{attribute 'pack_mode' := '1'} 
// ------------------------------------------------------------------------- 
//  SRCI Robot Library                                                
// ------------------------------------------------------------------------- 
//                                                                           
//  Object:      TelegramPlcToRobCyclicData                                       
//  Author:      Thorsten Brach                                                
//  Date:        2024-11-30
//
//  Description:                                              
//   
//                                                                           
//  Copyright: 
//    (C) 2024 Thorsten Brach. All rights reserved                                                                                                                                            
//             Licensed under the MIT License.
//                                                                           
//  Disclaimer:                                                                           
//    This project is provided without any guarantee and can be used for   
//    private and commercial purposes. Any use is at the user’s 
//    own risk and responsibility.
//
// -------------------------------------------------------------------------
TYPE TelegramPlcToRobCyclicData :
STRUCT
  /// Current Tool
  ToolNo  : BYTE;
  /// Current Frame
  FrameNo : BYTE;      
END_STRUCT
END_TYPE

{attribute 'pack_mode' := '1'} 
// ------------------------------------------------------------------------- 
//  SRCI Robot Library                                                
// ------------------------------------------------------------------------- 
//                                                                           
//  Object:      TelegramPlcToRobCyclicOptionalCartesianPos                                       
//  Author:      Thorsten Brach                                                
//  Date:        2024-06-01
//
//  Description:                                              
//   
//                                                                           
//  Copyright: 
//    (C) 2024 Thorsten Brach. All rights reserved                                                                                                                                            
//             Licensed under the MIT License.
//                                                                           
//  Disclaimer:                                                                           
//    This project is provided without any guarantee and can be used for   
//    private and commercial purposes. Any use is at the user’s 
//    own risk and responsibility.
//
// -------------------------------------------------------------------------
TYPE TelegramPlcToRobCyclicOptionalCartesianPosition :
STRUCT
  /// TCP Position on the X-Axis
  X           : REAL;
  /// TCP Position on the Y-Axis
  Y           : REAL;
  /// TCP Position on the Z-Axis
  Z           : REAL;
  /// Rotation around the X-Axis (RX)
  Rx          : REAL;
  /// Rotation around the Y-Axis (RY)
  Ry          : REAL;
  /// Rotation around the Z-Axis (RZ)
  Rz          : REAL;
  /// Configuration
  Config      : WORD;
  /// Turns of J1 and J2
  Turns_J2_J1 : BYTE;
  /// Turns of J3 and J4
  Turns_J4_J3 : BYTE;
  /// Turns of J6 and J5
  Turns_J6_J5 : BYTE;
  /// Turns of E1
  Turns_E1    : BYTE;
  /// Position of first external axis
  E1          : REAL;
END_STRUCT
END_TYPE

{attribute 'pack_mode' := '1'} 
// ------------------------------------------------------------------------- 
//  SRCI Robot Library                                                
// ------------------------------------------------------------------------- 
//                                                                           
//  Object:      TelegramPlcToRobCyclicOptionalCartesianPositionExt                                       
//  Author:      Thorsten Brach                                                
//  Date:        2024-06-01
//
//  Description:                                              
//   
//                                                                           
//  Copyright: 
//    (C) 2024 Thorsten Brach. All rights reserved                                                                                                                                            
//             Licensed under the MIT License.
//                                                                           
//  Disclaimer:                                                                           
//    This project is provided without any guarantee and can be used for   
//    private and commercial purposes. Any use is at the user’s 
//    own risk and responsibility.
//
// -------------------------------------------------------------------------
TYPE TelegramPlcToRobCyclicOptionalCartesianPositionExt :
STRUCT
  /// Position of second external axis
  E2 : REAL;
  /// Position of third external axis
  E3 : REAL;
  /// Position of fourth external axis
  E4 : REAL;
  /// Position of fifth external axis
  E5 : REAL;
  /// Position of sixth external axis
  E6 : REAL;    
END_STRUCT
END_TYPE

{attribute 'pack_mode' := '1'} 
// ------------------------------------------------------------------------- 
//  SRCI Robot Library                                                
// ------------------------------------------------------------------------- 
//                                                                           
//  Object:      TelegramPlcToRobCyclicOptionalCurrent                                       
//  Author:      Thorsten Brach                                                
//  Date:        2024-06-01
//
//  Description:                                              
//   
//                                                                           
//  Copyright: 
//    (C) 2024 Thorsten Brach. All rights reserved                                                                                                                                            
//             Licensed under the MIT License.
//                                                                           
//  Disclaimer:                                                                           
//    This project is provided without any guarantee and can be used for   
//    private and commercial purposes. Any use is at the user’s 
//    own risk and responsibility.
//
// -------------------------------------------------------------------------
TYPE TelegramPlcToRobCyclicOptionalCurrent :
STRUCT
  /// Current of first joint of the robot
  J1 : REAL;
  /// Current of second joint of the robot
  J2 : REAL;
  /// Current of third joint of the robot
  J3 : REAL;
  /// Current of fourth joint of the robot
  J4 : REAL;
  /// Current of fifth joint of the robot
  J5 : REAL;
  /// Current of sixth joint of the robot
  J6 : REAL;  
END_STRUCT
END_TYPE

{attribute 'pack_mode' := '1'} 
// ------------------------------------------------------------------------- 
//  SRCI Robot Library                                                
// ------------------------------------------------------------------------- 
//                                                                           
//  Object:      TelegramPlcToRobCyclicOptionalCurrentExt                                       
//  Author:      Thorsten Brach                                                
//  Date:        2024-06-01
//
//  Description:                                              
//   
//                                                                           
//  Copyright: 
//    (C) 2024 Thorsten Brach. All rights reserved                                                                                                                                            
//             Licensed under the MIT License.
//                                                                           
//  Disclaimer:                                                                           
//    This project is provided without any guarantee and can be used for   
//    private and commercial purposes. Any use is at the user’s 
//    own risk and responsibility.
//
// -------------------------------------------------------------------------
TYPE TelegramPlcToRobCyclicOptionalCurrentExt :
STRUCT
  /// Current of first external joint of the robot
  E1 : REAL;
  /// Current of second external axis
  E2: REAL;
  /// Current of third external axis
  E3: REAL;
  /// Current of fourth external axis
  E4: REAL;
  /// Current of fifth external axis
  E5: REAL;
  /// Current of sixth external axis
  E6: REAL;  
END_STRUCT
END_TYPE

{attribute 'pack_mode' := '1'} 
// ------------------------------------------------------------------------- 
//  SRCI Robot Library                                                
// ------------------------------------------------------------------------- 
//                                                                           
//  Object:      TelegramPlcToRobCyclicOptionalForce                                       
//  Author:      Thorsten Brach                                                
//  Date:        2024-06-01
//
//  Description:                                              
//   
//                                                                           
//  Copyright: 
//    (C) 2024 Thorsten Brach. All rights reserved                                                                                                                                            
//             Licensed under the MIT License.
//                                                                           
//  Disclaimer:                                                                           
//    This project is provided without any guarantee and can be used for   
//    private and commercial purposes. Any use is at the user’s 
//    own risk and responsibility.
//
// -------------------------------------------------------------------------
TYPE TelegramPlcToRobCyclicOptionalForce :
STRUCT
  /// Force on the X-Axis
  X : REAL;
  /// Force on the Y-Axis
  Y : REAL;
  /// Force on the Z-Axis
  Z : REAL;
  /// Force around the X-Axis (RX)
  Rx : REAL;
  /// Force around the Y-Axis (RY)
  Ry : REAL;
  /// Force around the Z-Axis (RZ)
  Rz : REAL;
END_STRUCT
END_TYPE

{attribute 'pack_mode' := '1'} 
// ------------------------------------------------------------------------- 
//  SRCI Robot Library                                                
// ------------------------------------------------------------------------- 
//                                                                           
//  Object:      TelegramPlcToRobCyclicOptionalForceExt                                       
//  Author:      Thorsten Brach                                                
//  Date:        2024-06-01
//
//  Description:                                              
//   
//                                                                           
//  Copyright: 
//    (C) 2024 Thorsten Brach. All rights reserved                                                                                                                                            
//             Licensed under the MIT License.
//                                                                           
//  Disclaimer:                                                                           
//    This project is provided without any guarantee and can be used for   
//    private and commercial purposes. Any use is at the user’s 
//    own risk and responsibility.
//
// -------------------------------------------------------------------------
TYPE TelegramPlcToRobCyclicOptionalForceExt :
STRUCT
  /// Force on the external axis 1
  E1 : REAL;
  /// Force on the external axis 2
  E2 : REAL;
  /// Force on the external axis 3
  E3 : REAL;
  /// Force om the external axis 4
  E4 : REAL;
  /// Force on the external axis 5
  E5 : REAL;
  /// Force on the external axis 6
  E6 : REAL;
END_STRUCT
END_TYPE

{attribute 'pack_mode' := '1'} 
// ------------------------------------------------------------------------- 
//  SRCI Robot Library                                                
// ------------------------------------------------------------------------- 
//                                                                           
//  Object:      TelegramPlcToRobCyclicOptionalJointPosition                                       
//  Author:      Thorsten Brach                                                
//  Date:        2024-06-01
//
//  Description:                                              
//   
//                                                                           
//  Copyright: 
//    (C) 2024 Thorsten Brach. All rights reserved                                                                                                                                            
//             Licensed under the MIT License.
//                                                                           
//  Disclaimer:                                                                           
//    This project is provided without any guarantee and can be used for   
//    private and commercial purposes. Any use is at the user’s 
//    own risk and responsibility.
//
// -------------------------------------------------------------------------
TYPE TelegramPlcToRobCyclicOptionalJointPosition :
STRUCT
  /// Position of first joint of the robot
  J1 : REAL;
  /// Position of second joint of the robot
  J2 : REAL;
  /// Position of third joint of the robot
  J3 : REAL;
  /// Position of fourth joint of the robot
  J4 : REAL;
  /// Position of fifth joint of the robot
  J5 : REAL;
  /// Position of sixth joint of the robot
  J6 : REAL;
  /// Position of first external axis 
  E1 : REAL;  
END_STRUCT
END_TYPE

{attribute 'pack_mode' := '1'} 
// ------------------------------------------------------------------------- 
//  SRCI Robot Library                                                
// ------------------------------------------------------------------------- 
//                                                                           
//  Object:      TelegramPlcToRobCyclicOptionalJointPositionExt                                       
//  Author:      Thorsten Brach                                                
//  Date:        2024-06-01
//
//  Description:                                              
//   
//                                                                           
//  Copyright: 
//    (C) 2024 Thorsten Brach. All rights reserved                                                                                                                                            
//             Licensed under the MIT License.
//                                                                           
//  Disclaimer:                                                                           
//    This project is provided without any guarantee and can be used for   
//    private and commercial purposes. Any use is at the user’s 
//    own risk and responsibility.
//
// -------------------------------------------------------------------------
TYPE TelegramPlcToRobCyclicOptionalJointPositionExt :
STRUCT
  /// Position of second external axis
  E2: REAL;
  /// Position of third external axis
  E3: REAL;
  /// Position of fourth external axis
  E4: REAL;
  /// Position of fifth external axis
  E5: REAL;
  /// Position of sixth external axis
  E6: REAL;    
END_STRUCT
END_TYPE

{attribute 'pack_mode' := '1'} 
// ------------------------------------------------------------------------- 
//  SRCI Robot Library                                                
// ------------------------------------------------------------------------- 
//                                                                           
//  Object:      TelegramPlcToRobCyclicOptionalSubProgramData                                       
//  Author:      Thorsten Brach                                                
//  Date:        2024-06-01
//
//  Description:                                              
//   
//                                                                           
//  Copyright: 
//    (C) 2024 Thorsten Brach. All rights reserved                                                                                                                                            
//             Licensed under the MIT License.
//                                                                           
//  Disclaimer:                                                                           
//    This project is provided without any guarantee and can be used for   
//    private and commercial purposes. Any use is at the user’s 
//    own risk and responsibility.
//
// -------------------------------------------------------------------------
TYPE TelegramPlcToRobCyclicOptionalSubProgramData :
STRUCT
  /// Sub program data
  /// ST-FIX F179: size from RobotLibraryConstants.CYCLIC_SUB_PROGRAM_DATA_MAX
  Data : ARRAY [0..RobotLibraryConstants.CYCLIC_SUB_PROGRAM_DATA_MAX] OF BYTE;
END_STRUCT
END_TYPE

{attribute 'pack_mode' := '1'} 
// ------------------------------------------------------------------------- 
//  SRCI Robot Library                                                
// ------------------------------------------------------------------------- 
//                                                                           
//  Object:      TelegramPlcToRobCyclicOptionalData                                       
//  Author:      Thorsten Brach                                                
//  Date:        2024-06-01
//
//  Description:                                              
//   
//                                                                           
//  Copyright: 
//    (C) 2024 Thorsten Brach. All rights reserved                                                                                                                                            
//             Licensed under the MIT License.
//                                                                           
//  Disclaimer:                                                                           
//    This project is provided without any guarantee and can be used for   
//    private and commercial purposes. Any use is at the user’s 
//    own risk and responsibility.
//
// -------------------------------------------------------------------------
TYPE TelegramPlcToRobCyclicOptionalData :
STRUCT
  /// Transmit cyclic data from PLC to RC for the usage in a subprogram on the RC called via the function “CallSubprogram”
  SubProgramData        :  TelegramPlcToRobCyclicOptionalSubProgramData;
  /// short cartesian position with TCP position (X, Y,Z), rotation (RX, RY, RZ), configuration bytes (Config, TurnNumber), position of first external axis (E1) and corresponding coordinate systems (ToolNo, FrameNo)
  CartesianPosition     :  TelegramPlcToRobCyclicOptionalCartesianPosition;
  /// the external axis values for an extended cartesian position (E2, E3, E4, E5, E6) 
  /// When selected, Tool and Frame will automatically cyclically be sent from client to server.
  CartesianPositionExt  :  TelegramPlcToRobCyclicOptionalCartesianPositionExt;
  /// short axes position with joint values (J1, J2, J3,J4, J5, J6) and position of first external axis (E1)
  JointPosition         :  TelegramPlcToRobCyclicOptionalJointPosition;
  /// the external axis values for an extended joint position (E2, E3, E4, E5, E6)
  JointPositionExt      :  TelegramPlcToRobCyclicOptionalJointPositionExt;
  /// force with the divided forces in the individual directions (X, Y, Z, RX, RY, RZ)
  Force                 :  TelegramPlcToRobCyclicOptionalForce;
  /// current force for the external axis (E1, E2, E3, E4, E5, E6)
  ForceExt              :  TelegramPlcToRobCyclicOptionalForceExt;
  /// ctual axes current of individual axes (J1, J2, J3, J4, J5, J6)
  Current               :  TelegramPlcToRobCyclicOptionalCurrent;
  /// actual current for the external axis (E1, E2,E3, E4, E5, E6)
  CurrentExt            :  TelegramPlcToRobCyclicOptionalCurrentExt;
END_STRUCT
END_TYPE

{attribute 'pack_mode' := '1'} 
// ------------------------------------------------------------------------- 
//  SRCI Robot Library                                                
// ------------------------------------------------------------------------- 
//                                                                           
//  Object:      TelegramPlcToRobFooter                                       
//  Author:      Thorsten Brach                                                
//  Date:        2024-06-01
//
//  Description:                                              
//   
//                                                                           
//  Copyright: 
//    (C) 2024 Thorsten Brach. All rights reserved                                                                                                                                            
//             Licensed under the MIT License.
//                                                                           
//  Disclaimer:                                                                           
//    This project is provided without any guarantee and can be used for   
//    private and commercial purposes. Any use is at the user’s 
//    own risk and responsibility.
//
// -------------------------------------------------------------------------
TYPE TelegramPlcToRobFooter :
STRUCT
  /// Life Sign
  LifeSign : BYTE;
  /// Reserve
  Reserve  : BYTE;
END_STRUCT
END_TYPE

{attribute 'pack_mode' := '1'} 
// ------------------------------------------------------------------------- 
//  SRCI Robot Library                                                
// ------------------------------------------------------------------------- 
//                                                                           
//  Object:      TelegramPlcToRobFragment                                       
//  Author:      Thorsten Brach                                                
//  Date:        2024-06-01
//
//  Description:                                              
//   
//                                                                           
//  Copyright: 
//    (C) 2024 Thorsten Brach. All rights reserved                                                                                                                                            
//             Licensed under the MIT License.
//                                                                           
//  Disclaimer:                                                                           
//    This project is provided without any guarantee and can be used for   
//    private and commercial purposes. Any use is at the user’s 
//    own risk and responsibility.
//
// -------------------------------------------------------------------------
TYPE TelegramPlcToRobFragment :
STRUCT
  /// Header
  Header  : TelegramPlcToRobFragmentHeader;
  /// Command
  Command : TelegramPlcToRobCommand;
END_STRUCT
END_TYPE

{attribute 'pack_mode' := '1'} 
// ------------------------------------------------------------------------- 
//  SRCI Robot Library                                                
// ------------------------------------------------------------------------- 
//                                                                           
//  Object:      TelegramPlcToRobFragmentHeader                                       
//  Author:      Thorsten Brach                                                
//  Date:        2024-06-01
//
//  Description:                                              
//   
//                                                                           
//  Copyright: 
//    (C) 2024 Thorsten Brach. All rights reserved                                                                                                                                            
//             Licensed under the MIT License.
//                                                                           
//  Disclaimer:                                                                           
//    This project is provided without any guarantee and can be used for   
//    private and commercial purposes. Any use is at the user’s 
//    own risk and responsibility.
//
// -------------------------------------------------------------------------
TYPE TelegramPlcToRobFragmentHeader :
STRUCT
  /// Command Instance Identifier used to assign the CMD payload to a specific CMD instance
  CmdID          : UINT;
  /// Empty reserve byte
  Reserve        : BYTE;
  /// Fragment Action Byte
  FragmentAction : BYTE;
  /// Append received payload in the receive buffer at this position
  PayloadPointer : UINT;
  /// Length of the CMD payload
  PayloadLength  : UINT;  
END_STRUCT
END_TYPE

{attribute 'pack_mode' := '1'} 
// ------------------------------------------------------------------------- 
//  SRCI Robot Library                                                
// ------------------------------------------------------------------------- 
//                                                                           
//  Object:      TelegramPlcToRobHeader                                       
//  Author:      Thorsten Brach                                                
//  Date:        2024-06-01
//
//  Description:                                              
//   
//                                                                           
//  Copyright: 
//    (C) 2024 Thorsten Brach. All rights reserved                                                                                                                                            
//             Licensed under the MIT License.
//                                                                           
//  Disclaimer:                                                                           
//    This project is provided without any guarantee and can be used for   
//    private and commercial purposes. Any use is at the user’s 
//    own risk and responsibility.
//
// -------------------------------------------------------------------------
TYPE TelegramPlcToRobHeader :
STRUCT
  /// Version of SRCI specification
  /// Bit 0-4 : Minor version = Features        (0..31)
  /// Bit 5-7 : Major version = Breaking change (0..07)
  SRCIVersion            : BYTE;
  /// Fast stop trigger | LifeSign
  FastStop_LifeSign      : BYTE;
  /// Number of Bytes of the frame to be used for the telegram of the given Axisgroup. Direction client to server
  TelegramLengthPlcToRob : UINT;
  /// Number of Bytes of the frame to be used for the telegram of the given Axisgroup. Direction server to client
  TelegramLengthRobToPlc : UINT;
  /// Control AxesGroupID | Telegtam state control
  AxesGroupID_Control    : BYTE;
  /// Reserved for later versions
  Reserved               : BYTE;
  /// Configuration of the optional cyclic data. Direction client to server
  TelegramNumberPlcToRob : UINT;
  /// Configuration of the optional cyclic data. Direction server to client
  TelegramNumberRobToPlc : UINT;
  /// Date of the client in the format days since 1990.01.01
  ClientDate             : IEC_DATE;
  /// Time in the clients time zone in the format milliseconds since start of day
  ClientTime             : IEC_TIME;  
END_STRUCT
END_TYPE

{attribute 'pack_mode' := '1'} 
// ------------------------------------------------------------------------- 
//  SRCI Robot Library                                                
// ------------------------------------------------------------------------- 
//                                                                           
//  Object:      TelegramPlcToRobSequence                                       
//  Author:      Thorsten Brach                                                
//  Date:        2024-06-01
//
//  Description:                                              
//   
//                                                                           
//  Copyright: 
//    (C) 2024 Thorsten Brach. All rights reserved                                                                                                                                            
//             Licensed under the MIT License.
//                                                                           
//  Disclaimer:                                                                           
//    This project is provided without any guarantee and can be used for   
//    private and commercial purposes. Any use is at the user’s 
//    own risk and responsibility.
//
// -------------------------------------------------------------------------
TYPE TelegramPlcToRobSequence :
STRUCT
  /// Header
  Header   : TelegramPlcTorobSequenceHeader;
  /// Fragment
  Fragment : ARRAY[0..RobotLibraryParameter.FRAGMENT_MAX] OF TelegramPlcToRobFragment;
END_STRUCT
END_TYPE

{attribute 'pack_mode' := '1'} 
// ------------------------------------------------------------------------- 
//  SRCI Robot Library                                                
// ------------------------------------------------------------------------- 
//                                                                           
//  Object:      TelegramPlcTorobSequenceHeader                                       
//  Author:      Thorsten Brach                                                
//  Date:        2024-06-01
//
//  Description:                                              
//   
//                                                                           
//  Copyright: 
//    (C) 2024 Thorsten Brach. All rights reserved                                                                                                                                            
//             Licensed under the MIT License.
//                                                                           
//  Disclaimer:                                                                           
//    This project is provided without any guarantee and can be used for   
//    private and commercial purposes. Any use is at the user’s 
//    own risk and responsibility.
//
// -------------------------------------------------------------------------
TYPE TelegramPlcToRobSequenceHeader :
STRUCT
  /// Telegram Sequence and Acknowledgement number
  SEQ_ACK       : UINT;
  /// Length of the Telegram Sequence excluding this Telegram Sequence Header
  PayloadLength : UINT;
END_STRUCT
END_TYPE

{attribute 'pack_mode' := '1'} 
// ------------------------------------------------------------------------- 
//  SRCI Robot Library                                                
// ------------------------------------------------------------------------- 
//                                                                           
//  Object:      TelegramPlcToRob                                       
//  Author:      Thorsten Brach                                                
//  Date:        2024-06-01
//
//  Description:                                              
//   
//                                                                           
//  Copyright: 
//    (C) 2024 Thorsten Brach. All rights reserved                                                                                                                                            
//             Licensed under the MIT License.
//                                                                           
//  Disclaimer:                                                                           
//    This project is provided without any guarantee and can be used for   
//    private and commercial purposes. Any use is at the user’s 
//    own risk and responsibility.
//
// -------------------------------------------------------------------------
TYPE TelegramPlcToRob :
STRUCT
  /// Header
  Header         : TelegramPlcToRobHeader;
  /// Cyclic optional data
  Cyclic         : TelegramPlcToRobCyclicData;
  /// Cyclic optional data
  CyclicOptional : TelegramPlcToRobCyclicOptionalData;
  /// Sequence Data
  Sequence       : ARRAY[0..1] OF TelegramPlcToRobSequence;
  /// Footer
  Footer         : TelegramPlcToRobFooter;
END_STRUCT
END_TYPE

{attribute 'pack_mode' := '1'} 
// ------------------------------------------------------------------------- 
//  SRCI Robot Library                                                
// ------------------------------------------------------------------------- 
//                                                                           
//  Object:      TelegramPlcToRobMessage                                       
//  Author:      Thorsten Brach                                                
//  Date:        2024-11-02
//
//  Description:                                              
//   
//                                                                           
//  Copyright: 
//    (C) 2024 Thorsten Brach. All rights reserved                                                                                                                                            
//             Licensed under the MIT License.
//                                                                           
//  Disclaimer:                                                                           
//    This project is provided without any guarantee and can be used for   
//    private and commercial purposes. Any use is at the user’s 
//    own risk and responsibility.
//
// -------------------------------------------------------------------------
TYPE TelegramRobToPlcCommand :
STRUCT
  /// Header
  Header  : TelegramRobToPlcCommandHeader;
  /// Payload
  Payload : ARRAY[0..RobotLibraryParameter.RESPONSE_PAYLOAD_MAX] OF BYTE; 
END_STRUCT
END_TYPE

{attribute 'pack_mode' := '1'} 
// ------------------------------------------------------------------------- 
//  SRCI Robot Library                                                
// ------------------------------------------------------------------------- 
//                                                                           
//  Object:      TelegramPlcToRobMessageHeader                                       
//  Author:      Thorsten Brach                                                
//  Date:        2024-11-02
//
//  Description:                                              
//   
//                                                                           
//  Copyright: 
//    (C) 2024 Thorsten Brach. All rights reserved                                                                                                                                            
//             Licensed under the MIT License.
//                                                                           
//  Disclaimer:                                                                           
//    This project is provided without any guarantee and can be used for   
//    private and commercial purposes. Any use is at the user’s 
//    own risk and responsibility.
//
// -------------------------------------------------------------------------
TYPE TelegramRobToPlcCommandHeader :
STRUCT
  /// Parameter squence
  ParSeq               : BYTE;
  /// message Staet
  State                : CmdMessageState;
  /// Alarm Message Severity
  AlarmMessageSeverity : SINT;
  /// Alarm Message Code
  AlarmMessageCode     : UINT;
END_STRUCT
END_TYPE

{attribute 'pack_mode' := '1'} 
// ------------------------------------------------------------------------- 
//  SRCI Robot Library                                                
// ------------------------------------------------------------------------- 
//                                                                           
//  Object:      TelegramRobToPlcCyclicOptionalCartesianPosition                                       
//  Author:      Thorsten Brach                                                
//  Date:        2024-06-01
//
//  Description:                                              
//   
//                                                                           
//  Copyright: 
//    (C) 2024 Thorsten Brach. All rights reserved                                                                                                                                            
//             Licensed under the MIT License.
//                                                                           
//  Disclaimer:                                                                           
//    This project is provided without any guarantee and can be used for   
//    private and commercial purposes. Any use is at the user’s 
//    own risk and responsibility.
//
// -------------------------------------------------------------------------
TYPE TelegramRobToPlcCyclicOptionalCartesianPosition :
STRUCT
  /// TCP Position on the X-Axis
  X                    : REAL;
  /// TCP Position on the Y-Axis
  Y                    : REAL;
  /// TCP Position on the Z-Axis
  Z                    : REAL;
  /// Rotation around the X-Axis (RX)
  Rx                   : REAL;
  /// Rotation around the Y-Axis (RY)
  Ry                   : REAL;
  /// Rotation around the Z-Axis (RZ)
  Rz                   : REAL;
  /// Configuration
  Config               : WORD;
  /// Turns of J1 and J2
  Turns_J2_J1          : BYTE;
  /// Turns of J3 and J4
  Turns_J4_J3          : BYTE;
  /// Turns of J6 and J5
  Turns_J6_J5          : BYTE;
  /// Turns of E1
  Turns_E1             : BYTE;
  /// Position of first external axis
  E1                   : REAL;  
  /// Tool Number
  ToolNo               : USINT;
  /// Frane Number
  FrameNo              : USINT;
  /// Currently used tool number
  CurrentlyUsedToolNo  : USINT;
  /// Currently used frame number
  CurrentlyUsedFrameNo : USINT;
  /// Reserve
  Reserve_1            : BYTE;
  /// Reserve
  Reserve_2            : BYTE;  
END_STRUCT
END_TYPE

{attribute 'pack_mode' := '1'} 
// ------------------------------------------------------------------------- 
//  SRCI Robot Library                                                
// ------------------------------------------------------------------------- 
//                                                                           
//  Object:      TelegramRobToPlcCyclicOptionalCartesianPosExt                                       
//  Author:      Thorsten Brach                                                
//  Date:        2024-06-01
//
//  Description:                                              
//   
//                                                                           
//  Copyright: 
//    (C) 2024 Thorsten Brach. All rights reserved                                                                                                                                            
//             Licensed under the MIT License.
//                                                                           
//  Disclaimer:                                                                           
//    This project is provided without any guarantee and can be used for   
//    private and commercial purposes. Any use is at the user’s 
//    own risk and responsibility.
//
// -------------------------------------------------------------------------
TYPE TelegramRobToPlcCyclicOptionalCartesianPositionExt :
STRUCT
  /// Position of second external axis
  E2 : REAL;
  /// Position of third external axis
  E3 : REAL;
  /// Position of fourth external axis
  E4 : REAL;
  /// Position of fifth external axis
  E5 : REAL;
  /// Position of sixth external axis
  E6 : REAL;    
END_STRUCT
END_TYPE

{attribute 'pack_mode' := '1'} 
// ------------------------------------------------------------------------- 
//  SRCI Robot Library                                                
// ------------------------------------------------------------------------- 
//                                                                           
//  Object:      TelegramRobToPlcCyclicOptionalCurrent                                       
//  Author:      Thorsten Brach                                                
//  Date:        2024-06-01
//
//  Description:                                              
//   
//                                                                           
//  Copyright: 
//    (C) 2024 Thorsten Brach. All rights reserved                                                                                                                                            
//             Licensed under the MIT License.
//                                                                           
//  Disclaimer:                                                                           
//    This project is provided without any guarantee and can be used for   
//    private and commercial purposes. Any use is at the user’s 
//    own risk and responsibility.
//
// -------------------------------------------------------------------------
TYPE TelegramRobToPlcCyclicOptionalCurrent :
STRUCT
  /// Current of first joint of the robot
  J1 : REAL;
  /// Current of second joint of the robot
  J2 : REAL;
  /// Current of third joint of the robot
  J3 : REAL;
  /// Current of fourth joint of the robot
  J4 : REAL;
  /// Current of fifth joint of the robot
  J5 : REAL;
  /// Current of sixth joint of the robot
  J6 : REAL;  
END_STRUCT
END_TYPE

{attribute 'pack_mode' := '1'} 
// ------------------------------------------------------------------------- 
//  SRCI Robot Library                                                
// ------------------------------------------------------------------------- 
//                                                                           
//  Object:      TelegramRobToPlcCyclicOptionalCurrentExt                                       
//  Author:      Thorsten Brach                                                
//  Date:        2024-06-01
//
//  Description:                                              
//   
//                                                                           
//  Copyright: 
//    (C) 2024 Thorsten Brach. All rights reserved                                                                                                                                            
//             Licensed under the MIT License.
//                                                                           
//  Disclaimer:                                                                           
//    This project is provided without any guarantee and can be used for   
//    private and commercial purposes. Any use is at the user’s 
//    own risk and responsibility.
//
// -------------------------------------------------------------------------
TYPE TelegramRobToPlcCyclicOptionalCurrentExt :
STRUCT
  /// Current of first external joint of the robot
  E1: REAL;
  /// Current of second external axis
  E2: REAL;
  /// Current of third external axis
  E3: REAL;
  /// Current of fourth external axis
  E4: REAL;
  /// Current of fifth external axis
  E5: REAL;
  /// Current of sixth external axis
  E6: REAL;  
END_STRUCT
END_TYPE

{attribute 'pack_mode' := '1'} 
// ------------------------------------------------------------------------- 
//  SRCI Robot Library                                                
// ------------------------------------------------------------------------- 
//                                                                           
//  Object:      TelegramRobToPlcCyclicOptionalForce                                       
//  Author:      Thorsten Brach                                                
//  Date:        2024-06-01
//
//  Description:                                              
//   
//                                                                           
//  Copyright: 
//    (C) 2024 Thorsten Brach. All rights reserved                                                                                                                                            
//             Licensed under the MIT License.
//                                                                           
//  Disclaimer:                                                                           
//    This project is provided without any guarantee and can be used for   
//    private and commercial purposes. Any use is at the user’s 
//    own risk and responsibility.
//
// -------------------------------------------------------------------------
TYPE TelegramRobToPlcCyclicOptionalForce :
STRUCT
  /// Force on the X-Axis
  X : REAL;
  /// Force on the Y-Axis
  Y : REAL;
  /// Force on the Z-Axis
  Z : REAL;
  /// Force around the X-Axis (RX)
  Rx : REAL;
  /// Force around the Y-Axis (RY)
  Ry : REAL;
  /// Force around the Z-Axis (RZ)
  Rz : REAL;
END_STRUCT
END_TYPE

{attribute 'pack_mode' := '1'} 
// ------------------------------------------------------------------------- 
//  SRCI Robot Library                                                
// ------------------------------------------------------------------------- 
//                                                                           
//  Object:      TelegramRobToPlcCyclicOptionalForceExt                                       
//  Author:      Thorsten Brach                                                
//  Date:        2024-06-01
//
//  Description:                                              
//   
//                                                                           
//  Copyright: 
//    (C) 2024 Thorsten Brach. All rights reserved                                                                                                                                            
//             Licensed under the MIT License.
//                                                                           
//  Disclaimer:                                                                           
//    This project is provided without any guarantee and can be used for   
//    private and commercial purposes. Any use is at the user’s 
//    own risk and responsibility.
//
// -------------------------------------------------------------------------
TYPE TelegramRobToPlcCyclicOptionalForceExt :
STRUCT
  /// Force on the external axis 1
  E1 : REAL;
  /// Force on the external axis 2
  E2 : REAL;
  /// Force on the external axis 3
  E3 : REAL;
  /// Force om the external axis 4
  E4 : REAL;
  /// Force on the external axis 5
  E5 : REAL;
  /// Force on the external axis 6
  E6 : REAL;
END_STRUCT
END_TYPE

{attribute 'pack_mode' := '1'} 
// ------------------------------------------------------------------------- 
//  SRCI Robot Library                                                
// ------------------------------------------------------------------------- 
//                                                                           
//  Object:      TelegramRobToPlcCyclicOptionalJointPosition                                       
//  Author:      Thorsten Brach                                                
//  Date:        2024-06-01
//
//  Description:                                              
//   
//                                                                           
//  Copyright: 
//    (C) 2024 Thorsten Brach. All rights reserved                                                                                                                                            
//             Licensed under the MIT License.
//                                                                           
//  Disclaimer:                                                                           
//    This project is provided without any guarantee and can be used for   
//    private and commercial purposes. Any use is at the user’s 
//    own risk and responsibility.
//
// -------------------------------------------------------------------------
TYPE TelegramRobToPlcCyclicOptionalJointPosition :
STRUCT
  /// Position of first joint of the robot
  J1 : REAL;
  /// Position of second joint of the robot
  J2 : REAL;
  /// Position of third joint of the robot
  J3 : REAL;
  /// Position of fourth joint of the robot
  J4 : REAL;
  /// Position of fifth joint of the robot
  J5 : REAL;
  /// Position of sixth joint of the robot
  J6 : REAL;
  /// Position of first external axis 
  E1 : REAL;  
  /// Reserve
  E1_Reserve : WORD;
END_STRUCT
END_TYPE

{attribute 'pack_mode' := '1'} 
// ------------------------------------------------------------------------- 
//  SRCI Robot Library                                                
// ------------------------------------------------------------------------- 
//                                                                           
//  Object:      TelegramRobToPlcCyclicOptionalJointPositionExt                                       
//  Author:      Thorsten Brach                                                
//  Date:        2024-06-01
//
//  Description:                                              
//   
//                                                                           
//  Copyright: 
//    (C) 2024 Thorsten Brach. All rights reserved                                                                                                                                            
//             Licensed under the MIT License.
//                                                                           
//  Disclaimer:                                                                           
//    This project is provided without any guarantee and can be used for   
//    private and commercial purposes. Any use is at the user’s 
//    own risk and responsibility.
//
// -------------------------------------------------------------------------
TYPE TelegramRobToPlcCyclicOptionalJointPositionExt :
STRUCT
  /// Position of second external axis
  E2: REAL;
  /// Position of third external axis
  E3: REAL;
  /// Position of fourth external axis
  E4: REAL;
  /// Position of fifth external axis
  E5: REAL;
  /// Position of sixth external axis
  E6: REAL;    
END_STRUCT
END_TYPE

{attribute 'pack_mode' := '1'} 
// ------------------------------------------------------------------------- 
//  SRCI Robot Library                                                
// ------------------------------------------------------------------------- 
//                                                                           
//  Object:      TelegramRobToPlcCyclicOptionalSubProgramData                                       
//  Author:      Thorsten Brach                                                
//  Date:        2024-06-01
//
//  Description:                                              
//   
//                                                                           
//  Copyright: 
//    (C) 2024 Thorsten Brach. All rights reserved                                                                                                                                            
//             Licensed under the MIT License.
//                                                                           
//  Disclaimer:                                                                           
//    This project is provided without any guarantee and can be used for   
//    private and commercial purposes. Any use is at the user’s 
//    own risk and responsibility.
//
// -------------------------------------------------------------------------
TYPE TelegramRobToPlcCyclicOptionalSubProgramData :
STRUCT
  /// Sub program data
  /// ST-FIX F179: size from RobotLibraryConstants.CYCLIC_SUB_PROGRAM_DATA_MAX (was 0..25 with a warning pragma)
  Data : ARRAY [0..RobotLibraryConstants.CYCLIC_SUB_PROGRAM_DATA_MAX] OF BYTE;
END_STRUCT
END_TYPE

{attribute 'pack_mode' := '1'} 
// ------------------------------------------------------------------------- 
//  SRCI Robot Library                                                
// ------------------------------------------------------------------------- 
//                                                                           
//  Object:      TelegramRobToPlcCyclicOptionalData                                       
//  Author:      Thorsten Brach                                                
//  Date:        2024-06-01
//
//  Description:                                              
//   
//                                                                           
//  Copyright: 
//    (C) 2024 Thorsten Brach. All rights reserved                                                                                                                                            
//             Licensed under the MIT License.
//                                                                           
//  Disclaimer:                                                                           
//    This project is provided without any guarantee and can be used for   
//    private and commercial purposes. Any use is at the user’s 
//    own risk and responsibility.
//
// -------------------------------------------------------------------------
TYPE TelegramRobToPlcCyclicOptionalData :
STRUCT
    /// Transmit cyclic data from PLC to RC for the usage in a subprogram on the RC called via the function “CallSubprogram”
  SubProgramData        :  TelegramRobToPlcCyclicOptionalSubProgramData;
  /// cartesian position with TCP position (X, Y,Z), rotation (RX, RY, RZ), configuration bytes (Config, TurnNumber), position of first external axis (E1) and corresponding coordinate systems (ToolNo, FrameNo)
  CartesianPosition     :  TelegramRobToPlcCyclicOptionalCartesianPosition;
  /// axes position with joint values (J1, J2, J3,J4, J5, J6) and position of first external axis (E1)
  JointPosition         :  TelegramRobToPlcCyclicOptionalJointPosition;
  /// force with the divided forces in the individual directions (X, Y, Z, RX, RY, RZ)
  Force                 :  TelegramRobToPlcCyclicOptionalForce;
  /// Transmit actual axes current of individual axes (J1, J2, J3, J4, J5, J6)
  Current               :  TelegramRobToPlcCyclicOptionalCurrent;
  /// Set to 1 to define two Sequences in one Telegram. If activated, 
  /// 2 sequences also has to be activated in the ClientServer direction.
  TwoSequences          : BYTE;  
  /// Transmit the external axis values for an extended cartesian position (E2, E3, E4, E5, E6)
  /// When selected, Tool and Frame will automatically cyclically be sent from client to server.
  CartesianPositionExt  :  TelegramRobToPlcCyclicOptionalCartesianPositionExt;
  /// Transmit the external axis values for an extended joint position (E2, E3, E4, E5, E6)
  JointPositionExt      :  TelegramRobToPlcCyclicOptionalJointPositionExt;
  /// Transmit actual axes force of individual axes (E1, E2, E3, E4, E5, E6)
  ForceExt              :  TelegramRobToPlcCyclicOptionalCurrentExt;
  /// Transmit actual axes current of individual axes (E1, E2, E3, E4, E5, E6)
  CurrentExt            :  TelegramRobToPlcCyclicOptionalCurrentExt;
END_STRUCT
END_TYPE

{attribute 'pack_mode' := '1'} 
// ------------------------------------------------------------------------- 
//  SRCI Robot Library                                                
// ------------------------------------------------------------------------- 
//                                                                           
//  Object:      TelegramPlcToRobFooter                                       
//  Author:      Thorsten Brach                                                
//  Date:        2024-06-01
//
//  Description:                                              
//   
//                                                                           
//  Copyright: 
//    (C) 2024 Thorsten Brach. All rights reserved                                                                                                                                            
//             Licensed under the MIT License.
//                                                                           
//  Disclaimer:                                                                           
//    This project is provided without any guarantee and can be used for   
//    private and commercial purposes. Any use is at the user’s 
//    own risk and responsibility.
//
// -------------------------------------------------------------------------
TYPE TelegramRobToPlcFooter :
STRUCT
  /// Reserve
  Reserve  : BYTE;
  /// Life Sign
  LifeSign : BYTE;
END_STRUCT
END_TYPE

{attribute 'pack_mode' := '1'} 
// ------------------------------------------------------------------------- 
//  SRCI Robot Library                                                
// ------------------------------------------------------------------------- 
//                                                                           
//  Object:      TelegramPlcToRobFragment                                       
//  Author:      Thorsten Brach                                                
//  Date:        2024-11-02
//
//  Description:                                              
//   
//                                                                           
//  Copyright: 
//    (C) 2024 Thorsten Brach. All rights reserved                                                                                                                                            
//             Licensed under the MIT License.
//                                                                           
//  Disclaimer:                                                                           
//    This project is provided without any guarantee and can be used for   
//    private and commercial purposes. Any use is at the user’s 
//    own risk and responsibility.
//
// -------------------------------------------------------------------------
TYPE TelegramRobToPlcFragment :
STRUCT
  /// Header
  Header  : TelegramRobToPlcFragmentHeader;
  /// Command
  Command : TelegramRobToPlcCommand;
END_STRUCT
END_TYPE

{attribute 'pack_mode' := '1'} 
// ------------------------------------------------------------------------- 
//  SRCI Robot Library                                                
// ------------------------------------------------------------------------- 
//                                                                           
//  Object:      TelegramPlcToRobFragmentHeader                                       
//  Author:      Thorsten Brach                                                
//  Date:        2024-11-02
//
//  Description:                                              
//   
//                                                                           
//  Copyright: 
//    (C) 2024 Thorsten Brach. All rights reserved                                                                                                                                            
//             Licensed under the MIT License.
//                                                                           
//  Disclaimer:                                                                           
//    This project is provided without any guarantee and can be used for   
//    private and commercial purposes. Any use is at the user’s 
//    own risk and responsibility.
//
// -------------------------------------------------------------------------
TYPE TelegramRobToPlcFragmentHeader :
STRUCT
  /// Command Instance Identifier used to assign the CMD payload to a specific CMD instance
  CmdID          : UINT;
  /// Empty reserve byte
  Reserve        : BYTE;
  /// Fragment Action Byte
  FragmentAction : BYTE;
  /// Append received payload in the receive buffer at this position
  PayloadPointer : UINT;
  /// Length of the CMD payload
  PayloadLength  : UINT;  
END_STRUCT
END_TYPE

{attribute 'pack_mode' := '1'} 
// ------------------------------------------------------------------------- 
//  SRCI Robot Library                                                
// ------------------------------------------------------------------------- 
//                                                                           
//  Object:      TelegramRobToPlcCyclic                                       
//  Author:      Thorsten Brach                                                
//  Date:        2024-06-01
//
//  Description:                                              
//   
//                                                                           
//  Copyright: 
//    (C) 2024 Thorsten Brach. All rights reserved                                                                                                                                            
//             Licensed under the MIT License.
//                                                                           
//  Disclaimer:                                                                           
//    This project is provided without any guarantee and can be used for   
//    private and commercial purposes. Any use is at the user’s 
//    own risk and responsibility.
//
// -------------------------------------------------------------------------
TYPE TelegramRobToPlcHeader :
STRUCT
  /// Version of SRCI specification
  /// Bit 0-4 : Minor version = Features        (0..31)
  /// Bit 5-7 : Major version = Breaking change (0..07)
  SRCIVersion   : VersionStruct;
  /// Connection alive signal
  LifeSign      : BYTE;
  /// Reserved byte
  Reserved      : BYTE;
  /// Initialization and Telegram control state
  TelegramState : TelegramState;
  /// Combination of various RA related states.
  StatusRobotArm: DWORD;
  /// Actual override in percentage encoding 
  Override      : UINT;
END_STRUCT
END_TYPE

{attribute 'pack_mode' := '1'} 
// ------------------------------------------------------------------------- 
//  SRCI Robot Library                                                
// ------------------------------------------------------------------------- 
//                                                                           
//  Object:      TelegramPlcToRobSequence                                       
//  Author:      Thorsten Brach                                                
//  Date:        2024-11-02
//
//  Description:                                              
//   
//                                                                           
//  Copyright: 
//    (C) 2024 Thorsten Brach. All rights reserved                                                                                                                                            
//             Licensed under the MIT License.
//                                                                           
//  Disclaimer:                                                                           
//    This project is provided without any guarantee and can be used for   
//    private and commercial purposes. Any use is at the user’s 
//    own risk and responsibility.
//
// -------------------------------------------------------------------------
TYPE TelegramRobToPlcSequence :
STRUCT
  /// Header
  Header   : TelegramRobToPlcSequenceHeader;
  /// Fragment
  Fragment : ARRAY[0..RobotLibraryParameter.FRAGMENT_MAX] OF TelegramRobToPlcFragment;
END_STRUCT
END_TYPE

{attribute 'pack_mode' := '1'} 
// ------------------------------------------------------------------------- 
//  SRCI Robot Library                                                
// ------------------------------------------------------------------------- 
//                                                                           
//  Object:      TelegramRobToPlcSequenceHeader                                       
//  Author:      Thorsten Brach                                                
//  Date:        2024-11-02
//
//  Description:                                              
//   
//                                                                           
//  Copyright: 
//    (C) 2024 Thorsten Brach. All rights reserved                                                                                                                                            
//             Licensed under the MIT License.
//                                                                           
//  Disclaimer:                                                                           
//    This project is provided without any guarantee and can be used for   
//    private and commercial purposes. Any use is at the user’s 
//    own risk and responsibility.
//
// -------------------------------------------------------------------------
TYPE TelegramRobToPlcSequenceHeader :
STRUCT
  /// Telegram Sequence and Acknowledgement number
  SEQ_ACK      : UINT;
  /// Length of the Telegram Sequence excluding this Telegram Sequence Header
  PayloadLength : UINT;
END_STRUCT
END_TYPE

{attribute 'pack_mode' := '1'} 
// ------------------------------------------------------------------------- 
//  SRCI Robot Library                                                
// ------------------------------------------------------------------------- 
//                                                                           
//  Object:      TelegramRobToPlc                                       
//  Author:      Thorsten Brach                                                
//  Date:        2024-06-01
//
//  Description:                                              
//   
//                                                                           
//  Copyright: 
//    (C) 2024 Thorsten Brach. All rights reserved                                                                                                                                            
//             Licensed under the MIT License.
//                                                                           
//  Disclaimer:                                                                           
//    This project is provided without any guarantee and can be used for   
//    private and commercial purposes. Any use is at the user’s 
//    own risk and responsibility.
//
// -------------------------------------------------------------------------
TYPE TelegramRobToPlc :
STRUCT
  /// Telegram Header
  Header               : TelegramRobToPlcHeader;
  /// Cyclic optional data
  CyclicOptional       : TelegramRobToPlcCyclicOptionalData;
  /// Sequence Data
  Sequence             : ARRAY[0..1] OF TelegramRobToPlcSequence;
  /// Footer
  Footer               : TelegramRobToPlcFooter;
END_STRUCT
END_TYPE

{attribute 'pack_mode' := '1'} 
// ------------------------------------------------------------------------- 
//  SRCI Robot Library                                                
// ------------------------------------------------------------------------- 
//                                                                           
//  Object:      Telegram                                       
//  Author:      Thorsten Brach                                                
//  Date:        2024-06-01
//
//  Description:                                              
//   
//                                                                           
//  Copyright: 
//    (C) 2024 Thorsten Brach. All rights reserved                                                                                                                                            
//             Licensed under the MIT License.
//                                                                           
//  Disclaimer:                                                                           
//    This project is provided without any guarantee and can be used for   
//    private and commercial purposes. Any use is at the user’s 
//    own risk and responsibility.
//
// -------------------------------------------------------------------------
TYPE Telegram :
STRUCT
  /// PLC to Robot
  PlcToRob : TelegramPlcToRob;
  /// Robot to PLC
  RobToPlc : TelegramRobToPlc;
END_STRUCT
END_TYPE

(* global variable list RobotLibraryConstants *)
{attribute 'qualified_only'}
// ------------------------------------------------------------------------- 
//  SRCI Robot Library                                                
// ------------------------------------------------------------------------- 
//                                                                           
//  Object:      RobotLibraryConstants                                       
//  Author:      Thorsten Brach                                                
//  Date:        2024-06-01
//
//  Description:                                              
//   
//                                                                           
//  Copyright: 
//    (C) 2024 Thorsten Brach. All rights reserved           
//             Licensed under the MIT License.                                                                                                                                 
//                                                                           
//  Disclaimer:                                                                           
//    This project is provided without any guarantee and can be used for   
//    private and commercial purposes. Any use is at the user’s 
//    own risk and responsibility.
//
// -------------------------------------------------------------------------
VAR_GLOBAL CONSTANT  
  /// Version of SRCI specification
  /// Bit 0-4 : Minor version = Features        (0..31)
  /// Bit 5-7 : Major version = Breaking change (0..07)
  SRCIVersion             : VersionStruct := ( MajorVersion := 1, MinorVersion := 5, PatchVersion := 0); // ST-FIX PLC library still says 1.3.0, but implements SRCI 1.5 (SDK: SRCI_VERSION 1.5)
  /// Version of the PLC library
  PLCLibraryVersion       : VersionStruct := ( MajorVersion := 1, MinorVersion := 5, PatchVersion := 7); // ST-FIX F166: the constant was not counted up (1.5.4 in library 1.5.5.0); now the release 1.5.7
  /// Minimal axes group ID
  AXES_GROUP_ID_MIN       : BYTE := 0;  
  /// Maximal axes groups ID
  AXES_GROUP_ID_MAX       : BYTE := 15;  
  /// OK = 0
  OK                      : DINT := 0;
  /// Running = 1
  RUNNING                 : DINT := 1;
  /// HasError = -1
  HAS_ERROR               : DINT := -1;  
  /// Null pointer
  XNULL                   : DWORD := 0;
  /// Null pointer
  NULL_POINTER            : POINTER TO BYTE := 0;
  /// Real conversion factor ( REAL * 100 -> TO_INT )
  REAL_CONVERSION_FACTOR  : REAL := 100;
  /// Active command
  ACTIVE_CMD              : UDINT := 1;
  /// Buffered command
  BUFFER_CMD              : UDINT := 2;
  /// Maximal length of additional text 
  MAX_ADD_TEXT_LENGTH     : DINT := 40;
  /// ST-FIX F108: characters of a log line per ReadServerLog response (SRCI SDK 1.1: 179;
  /// spec table 6-124: 187)
  SERVER_LOG_CONTENT_MAX  : DINT := 179;
  /// Upper index of the cyclic sub program data: 26 bytes (spec table 5-88, 6-711)
  /// ST-FIX F179: one constant for all arrays of the cyclic sub program data
  CYCLIC_SUB_PROGRAM_DATA_MAX : DINT := 25;
 END_VAR

(* global variable list RobotLibraryDefines *)
{attribute 'qualified_only'}
// ------------------------------------------------------------------------- 
//  SRCI Robot Library                                                
// ------------------------------------------------------------------------- 
//                                                                           
//  Object:      RobotLibraryDefines                                       
//  Author:      Thorsten Brach                                                
//  Date:        2024-06-01
//
//  Description:                                              
//   
//                                                                           
//  Copyright: 
//    (C) 2024 Thorsten Brach. All rights reserved           
//             Licensed under the MIT License.                                                                                                                                 
//                                                                           
//  Disclaimer:                                                                           
//    This project is provided without any guarantee and can be used for   
//    private and commercial purposes. Any use is at the user’s 
//    own risk and responsibility.
//
// -------------------------------------------------------------------------
VAR_GLOBAL
  /// Maximal length of type name
  MaxTypeNameLength  : INT;
END_VAR

(* global variable list RobotLibraryParameter *)
{attribute 'qualified_only'}
// ------------------------------------------------------------------------- 
//  SRCI Robot Library                                                
// ------------------------------------------------------------------------- 
//                                                                           
//  Object:      Parameter                                       
//  Author:      Thorsten Brach                                                
//  Date:        2024-06-01
//
//  Description:                                              
//   
//                                                                           
//  Copyright: 
//    (C) 2024 Thorsten Brach. All rights reserved                                                                                                                                            
//             Licensed under the MIT License.
//                                                                           
//  Disclaimer:                                                                           
//    This project is provided without any guarantee and can be used for   
//    private and commercial purposes. Any use is at the user’s 
//    own risk and responsibility.
//
// -------------------------------------------------------------------------
VAR_GLOBAL CONSTANT
  /// Maximal amount of tools
  /// SRCI_PLC_TEST: 20 like the SDK simulator (was the parameter of the library reference)
  TOOL_MAX                            : DINT := 20;
  /// Maximal amount of frames
  /// SRCI_PLC_TEST: 20 like the SDK simulator (was the parameter of the library reference)
  FRAME_MAX                           : DINT := 20;
  /// Maximal amount of loads
  /// SRCI_PLC_TEST: 20 like the SDK simulator (was the parameter of the library reference)
  LOAD_MAX                            : DINT := 20;  
  /// Maximal amount of work areas
  WORK_AREAS_MAX                      : DINT := 16;  
  /// Maximal amount of system logs
  SYSTEM_LOG_MAX                      : DINT := 32;  
  /// Maximal amount of message logs
  MESSAGE_LOG_MAX                     : DINT := 100;  
  /// Maximum string length for message texts
  MESSAGE_TEXT_LEN                    : DINT := 255;
  /// Maximal amount of List entries 
  LIST_ENTRIES_MAX                    : DINT := 100;
  /// Maximal amount of bytes for the parameter payload
  PARAMETER_PAYLOAD_MAX               : DINT := 255;  
  /// Maximal amount of bytes for the response payload
  RESPONSE_PAYLOAD_MAX                : DINT := 255;  
  /// Maximal amount of bytes that can be exchanged with the sub program on the RC
  SUB_PROGRAM_DATA_MAX                : DINT := 189;
  /// Maximal amount of spline data
  SPLINE_DATA_MAX                     : DINT := 64;
  /// Maximal amount of entries in the Active Command Register
  ACTIVE_CMD_REGISTER_ENTRIES_MAX     : DINT := 50;
  /// Maximal amount of message codes
  MESSAGE_CODES_MAX                   : DINT := 15;
  /// Maximal amount of fragments
  FRAGMENT_MAX                        : DINT := 31; // ST-FIX F52: 10 fragments (0..9) per telegram are too few - a 256 byte telegram holds up to 27 fragme
  /// Flag to indicate that the byte order must be changed
  SWAP_BYTE_ORDER                     : BOOL := TRUE; 
  /// Timeout for checking for invalid frames
  INVALID_FRAMES_CHECK_TIMEOUT        : TIME := T#60S;
  /// Warning limit for ACR registers running low
  ACR_USAGE_WARNING_LIMIT             : REAL := 80.0;  
  /// ST-FIX F108: maximal length of a log line of ReadServerLog / ReadClientLog (element of LogFile)
  LOG_LINE_LEN                        : DINT := 1023;
END_VAR

INTERFACE IMessageLogger
METHOD PUBLIC AddMessageLog
VAR_INPUT
  /// Message to add to the log
  MessageLog : AlarmMessage;
END_VAR
END_METHOD
METHOD PUBLIC AddSystemLog
VAR_INPUT
  /// System messafe to add to the log
  SystemLog : STRING(RobotLibraryParameter.MESSAGE_TEXT_LEN);
END_VAR
END_METHOD
END_INTERFACE

INTERFACE IRobotLibraryCommandFB
METHOD PUBLIC CallBack : DINT
VAR_INPUT
  /// Response data
  RspData : AxesGroupAcyclicAcrEntryRspBuffer;  
END_VAR
END_METHOD
PROPERTY CommandData : RobotLibrarySendDataFB
END_PROPERTY
END_INTERFACE

FUNCTION IsDefaultDynamicsEqual : BOOL
// ------------------------------------------------------------------------- 
//  SRCI Robot Library                                                
// ------------------------------------------------------------------------- 
//                                                                           
//  Object:      IsDefaultDynamicsEqual                                       
//  Author:      Thorsten Brach                                                
//  Date:        2025-04-23
//
//  Description:                                              
//   
//                                                                           
//  Copyright: 
//    (C) 2025 Thorsten Brach. All rights reserved                                                                                                                                            
//             Licensed under the MIT License.
//                                                                           
//  Disclaimer:                                                                           
//    This project is provided without any guarantee and can be used for   
//    private and commercial purposes. Any use is at the user’s 
//    own risk and responsibility.
//
// -------------------------------------------------------------------------
VAR_INPUT
  /// DefaultDynamics 1 to compare
  Data1           : DefaultDynamics;
  /// DefaultDynamics 2 to compare
  Data2           : DefaultDynamics;
  /// Flag to ignore the timestamp during the comparison
  IgnoreTimestamp : BOOL;
END_VAR

            IF (IgnoreTimestamp)
THEN
  Data1.Timestamp := Data2.Timestamp;
END_IF                    
                    
IsDefaultDynamicsEqual := ( SysDepMemCmp( pData1 := ADR(Data1), pData2 :=  ADR(Data2), DataLen := SIZEOF(Data1)) = RobotLibraryConstants.OK );
          
END_FUNCTION

FUNCTION IsFrameDataEqual : BOOL
// ------------------------------------------------------------------------- 
//  SRCI Robot Library                                                
// ------------------------------------------------------------------------- 
//                                                                           
//  Object:      IsFrameDataEqual                                       
//  Author:      Thorsten Brach                                                
//  Date:        2025-04-23
//
//  Description:                                              
//   
//                                                                           
//  Copyright: 
//    (C) 2025 Thorsten Brach. All rights reserved                                                                                                                                            
//             Licensed under the MIT License.
//                                                                           
//  Disclaimer:                                                                           
//    This project is provided without any guarantee and can be used for   
//    private and commercial purposes. Any use is at the user’s 
//    own risk and responsibility.
//
// -------------------------------------------------------------------------
VAR_INPUT
  /// FrameData 1 to compare
  Data1           : FrameData;
  /// FrameData 2 to compare
  Data2           : FrameData;
  /// Flag to ignore the timestamp during the comparison
  IgnoreTimestamp : BOOL;
END_VAR

            IF (IgnoreTimestamp)
THEN
  Data1.Timestamp := Data2.Timestamp;
END_IF                    
                    
IsFrameDataEqual := ( SysDepMemCmp( pData1 := ADR(Data1), pData2 :=  ADR(Data2), DataLen := SIZEOF(Data1)) = RobotLibraryConstants.OK );                    
          
END_FUNCTION

FUNCTION IsLoadDataEqual : BOOL
// ------------------------------------------------------------------------- 
//  SRCI Robot Library                                                
// ------------------------------------------------------------------------- 
//                                                                           
//  Object:      IsLoadDataEqual                                       
//  Author:      Thorsten Brach                                                
//  Date:        2025-04-23
//
//  Description:                                              
//   
//                                                                           
//  Copyright: 
//    (C) 2025 Thorsten Brach. All rights reserved                                                                                                                                            
//             Licensed under the MIT License.
//                                                                           
//  Disclaimer:                                                                           
//    This project is provided without any guarantee and can be used for   
//    private and commercial purposes. Any use is at the user’s 
//    own risk and responsibility.
//
// -------------------------------------------------------------------------
VAR_INPUT
  /// LoadData 1 to compare
  Data1           : LoadData;
  /// LoadData 2 to compare
  Data2           : LoadData;
  /// Flag to ignore the timestamp during the comparison
  IgnoreTimestamp : BOOL;
END_VAR

            IF (IgnoreTimestamp)
THEN
  Data1.Timestamp := Data2.Timestamp;
END_IF                    
                    
IsLoadDataEqual := ( SysDepMemCmp( pData1 := ADR(Data1), pData2 :=  ADR(Data2), DataLen := SIZEOF(Data1)) = RobotLibraryConstants.OK );
          
END_FUNCTION

FUNCTION IsReferenceDynamicsEqual : BOOL
// ------------------------------------------------------------------------- 
//  SRCI Robot Library                                                
// ------------------------------------------------------------------------- 
//                                                                           
//  Object:      IsReferenceDynamicsEqual                                       
//  Author:      Thorsten Brach                                                
//  Date:        2025-04-23
//
//  Description:                                              
//   
//                                                                           
//  Copyright: 
//    (C) 2025 Thorsten Brach. All rights reserved                                                                                                                                            
//             Licensed under the MIT License.
//                                                                           
//  Disclaimer:                                                                           
//    This project is provided without any guarantee and can be used for   
//    private and commercial purposes. Any use is at the user’s 
//    own risk and responsibility.
//
// -------------------------------------------------------------------------
VAR_INPUT
  /// ReferenceDynamics 1 to compare
  Data1           : ReferenceDynamics;
  /// ReferenceDynamics 2 to compare
  Data2           : ReferenceDynamics;
  /// Flag to ignore the timestamp during the comparison
  IgnoreTimestamp : BOOL;
END_VAR

            IF (IgnoreTimestamp)
THEN
  Data1.Timestamp := Data2.Timestamp;
END_IF                    
                    
IsReferenceDynamicsEqual := ( SysDepMemCmp( pData1 := ADR(Data1), pData2 :=  ADR(Data2), DataLen := SIZEOF(Data1)) = RobotLibraryConstants.OK );
          
END_FUNCTION

FUNCTION IsSwLimitsEqual : BOOL
// ------------------------------------------------------------------------- 
//  SRCI Robot Library                                                
// ------------------------------------------------------------------------- 
//                                                                           
//  Object:      IsSwLimitsEqual                                       
//  Author:      Thorsten Brach                                                
//  Date:        2025-04-23
//
//  Description:                                              
//   
//                                                                           
//  Copyright: 
//    (C) 2025 Thorsten Brach. All rights reserved                                                                                                                                            
//             Licensed under the MIT License.
//                                                                           
//  Disclaimer:                                                                           
//    This project is provided without any guarantee and can be used for   
//    private and commercial purposes. Any use is at the user’s 
//    own risk and responsibility.
//
// -------------------------------------------------------------------------
VAR_INPUT
  /// SW Limit 1 to compare
  Data1           : SWLimits;
  /// SW LIMIT 2 to compare
  Data2           : SWLimits;
  /// Flag to ignore the timestamp during the comparison
  IgnoreTimestamp : BOOL;
END_VAR

            IF (IgnoreTimestamp)
THEN
  Data1.Timestamp := Data2.Timestamp;
END_IF                    
                    
IsSwLimitsEqual := ( SysDepMemCmp( pData1 := ADR(Data1), pData2 :=  ADR(Data2), DataLen := SIZEOF(Data1)) = RobotLibraryConstants.OK );
          
END_FUNCTION

FUNCTION IsToolDataEqual : BOOL
// ------------------------------------------------------------------------- 
//  SRCI Robot Library                                                
// ------------------------------------------------------------------------- 
//                                                                           
//  Object:      IsToolDataEqual                                       
//  Author:      Thorsten Brach                                                
//  Date:        2025-04-23
//
//  Description:                                              
//   
//                                                                           
//  Copyright: 
//    (C) 2025 Thorsten Brach. All rights reserved                                                                                                                                            
//             Licensed under the MIT License.
//                                                                           
//  Disclaimer:                                                                           
//    This project is provided without any guarantee and can be used for   
//    private and commercial purposes. Any use is at the user’s 
//    own risk and responsibility.
//
// -------------------------------------------------------------------------
VAR_INPUT
  /// ToolData 1 to compare
  Data1           : ToolData;
  /// ToolData 2 to compare
  Data2           : ToolData;
  /// Flag to ignore the timestamp during the comparison
  IgnoreTimestamp : BOOL;
END_VAR

            IF (IgnoreTimestamp)
THEN
  Data1.Timestamp := Data2.Timestamp;
END_IF                    
                    
IsToolDataEqual := ( SysDepMemCmp( pData1 := ADR(Data1), pData2 :=  ADR(Data2), DataLen := SIZEOF(Data1)) = RobotLibraryConstants.OK );                    
          
END_FUNCTION

FUNCTION IsWorkAreaEqual : BOOL
// ------------------------------------------------------------------------- 
//  SRCI Robot Library                                                
// ------------------------------------------------------------------------- 
//                                                                           
//  Object:      IsWorkAreaEqual                                       
//  Author:      Thorsten Brach                                                
//  Date:        2025-04-23
//
//  Description:                                              
//   
//                                                                           
//  Copyright: 
//    (C) 2025 Thorsten Brach. All rights reserved                                                                                                                                            
//             Licensed under the MIT License.
//                                                                           
//  Disclaimer:                                                                           
//    This project is provided without any guarantee and can be used for   
//    private and commercial purposes. Any use is at the user’s 
//    own risk and responsibility.
//
// -------------------------------------------------------------------------
VAR_INPUT
  /// WorkArea 1 to compare
  Data1           : RobotWorkAreaData;
  /// WorkArea 2 to compare
  Data2           : RobotWorkAreaData;
  /// Flag to ignore the timestamp during the comparison
  IgnoreTimestamp : BOOL;
END_VAR

            IF (IgnoreTimestamp)
THEN
  Data1.Timestamp := Data2.Timestamp;
END_IF                    
                    
IsWorkAreaEqual := ( SysDepMemCmp( pData1 := ADR(Data1), pData2 :=  ADR(Data2), DataLen := SIZEOF(Data1)) = RobotLibraryConstants.OK );
          
END_FUNCTION

FUNCTION CheckTimeout : DINT
// ------------------------------------------------------------------------- 
//  SRCI Robot Library                                                
// ------------------------------------------------------------------------- 
//                                                                           
//  Object:      SwapBytes                                       
//  Author:      Thorsten Brach                                                
//  Date:        2024-12-18
//
//  Description:                                              
//   
//                                                                           
//  Copyright: 
//    (C) 2024 Thorsten Brach. All rights reserved                                                                                                                                            
//             Licensed under the MIT License.
//                                                                           
//  Disclaimer:                                                                           
//    This project is provided without any guarantee and can be used for   
//    private and commercial purposes. Any use is at the user’s 
//    own risk and responsibility.
//
// -------------------------------------------------------------------------
VAR_INPUT
  /// Reference to TON instance
  rTimer : REFERENCE TO TON;
END_VAR

            // Call timer 
rTimer();

// check if timer elapsed
IF (rTimer.Q = TRUE)
THEN
  // assign return value
  CheckTimeout := RobotLibraryConstants.OK;
ELSE
  // assign return value
  CheckTimeout := RobotLibraryConstants.RUNNING;
END_IF
          
END_FUNCTION

FUNCTION SetTimeout : DINT
// ------------------------------------------------------------------------- 
//  SRCI Robot Library                                                
// ------------------------------------------------------------------------- 
//                                                                           
//  Object:      SwapBytes                                       
//  Author:      Thorsten Brach                                                
//  Date:        2024-12-18
//
//  Description:                                              
//   
//                                                                           
//  Copyright: 
//    (C) 2024 Thorsten Brach. All rights reserved                                                                                                                                            
//             Licensed under the MIT License.
//                                                                           
//  Disclaimer:                                                                           
//    This project is provided without any guarantee and can be used for   
//    private and commercial purposes. Any use is at the user’s 
//    own risk and responsibility.
//
// -------------------------------------------------------------------------
VAR_INPUT
  /// Timeout to be set
  PT     : TIME;
  /// Reference to TON instance
  rTimer : REFERENCE TO TON;
END_VAR

            rTimer(IN := FALSE);          // Reset timer
rTimer(PT := PT, IN := TRUE); // Start timer

// assign return value
SetTimeout := RobotLibraryConstants.OK;
          
END_FUNCTION

FUNCTION DATE_TO_IEC_DATE : IEC_DATE
// ------------------------------------------------------------------------- 
//  SRCI Robot Library                                                
// ------------------------------------------------------------------------- 
//                                                                           
//  Object:      DATE_TO_IEC_DATE                                       
//  Author:      Thorsten Brach                                                
//  Date:        2024-06-01
//
//  Description:                                              
//   
//                                                                           
//  Copyright: 
//    (C) 2024 Thorsten Brach. All rights reserved                                                                                                                                            
//             Licensed under the MIT License.
//                                                                           
//  Disclaimer:                                                                           
//    This project is provided without any guarantee and can be used for   
//    private and commercial purposes. Any use is at the user’s 
//    own risk and responsibility.
//
// -------------------------------------------------------------------------
VAR_INPUT
  Value    : DATE;
END_VAR

VAR
 _tmpDate1 : DWORD;
 _tmpDate2 : DWORD;
 _initDate : DATE := DATE#1990-01-01;
 END_VAR

            // Siemens Dateformat is Day since 01.01.1990
// TwinCat Dateformat is seconds sinde 01.01.1970
// Calculation : 
// ( [TwinCat current date] - [ TwinCat 01.01.1970] ) / [Seconds a Day] = Days sinde 01.01.1990 (Siemens Format)

// copy date to dword
SysDepMemCpy( pDest := ADR(_tmpDate1), pSrc := ADR( Value   ), DataLen := SIZEOF( Value   ));
// copy date to dword
SysDepMemCpy( pDest := ADR(_tmpDate2), pSrc := ADR(_initDate), DataLen := SIZEOF(_initDate));

// calculate IEC Date :  
DATE_TO_IEC_DATE := UDINT_TO_UINT((_tmpDate1 - _tmpDate2) / 86400); // 86400 Seconds = 1 day 

          
END_FUNCTION

FUNCTION IEC_DATE_TO_DATE : DATE
// ------------------------------------------------------------------------- 
//  SRCI Robot Library                                                
// ------------------------------------------------------------------------- 
//                                                                           
//  Object:      IEC_DATE_TO_DATE                                       
//  Author:      Thorsten Brach                                                
//  Date:        2025-01-05
//
//  Description:                                              
//   
//                                                                           
//  Copyright: 
//    (C) 2025 Thorsten Brach. All rights reserved                                                                                                                                            
//             Licensed under the MIT License.
//                                                                           
//  Disclaimer:                                                                           
//    This project is provided without any guarantee and can be used for   
//    private and commercial purposes. Any use is at the user’s 
//    own risk and responsibility.
//
// -------------------------------------------------------------------------
VAR_INPUT
  Value    : IEC_DATE;
END_VAR

VAR
 _tmpDate1 : DWORD;
 _initDate : DATE := DATE#1990-01-01;
 END_VAR

            // Siemens Dateformat is Day since 01.01.1990
// TwinCat Dateformat is seconds sinde 01.01.1970
// Calculation : 
// ( [ TwinCat 01.01.1990] + [IEC Date]) * [Seconds a Day] = (TwinCat Format)

// copy date to dword
SysDepMemCpy( pDest := ADR(_tmpDate1), pSrc := ADR( _initDate ), DataLen := SIZEOF( _initDate ));

// calculate IEC Date :  
IEC_DATE_TO_DATE := DWORD_TO_DATE( _tmpDate1 + ( Value * 86400)); // 86400 Seconds = 1 day 
          
END_FUNCTION

FUNCTION IEC_TIME_TO_TIME : TOD
// ------------------------------------------------------------------------- 
//  SRCI Robot Library                                                
// ------------------------------------------------------------------------- 
//                                                                           
//  Object:      IEC_TIME_TO_TIME                                       
//  Author:      Thorsten Brach                                                
//  Date:        2025-01-05
//
//  Description:                                              
//   
//                                                                           
//  Copyright: 
//    (C) 2025 Thorsten Brach. All rights reserved                                                                                                                                            
//             Licensed under the MIT License.
//                                                                           
//  Disclaimer:                                                                           
//    This project is provided without any guarantee and can be used for   
//    private and commercial purposes. Any use is at the user’s 
//    own risk and responsibility.
//
// -------------------------------------------------------------------------
VAR_INPUT
  Value : IEC_TIME;
END_VAR

            IEC_TIME_TO_TIME := Value; 
          
END_FUNCTION

